Fanuc KAREL source: kt00010.KL

-- PROVISIONAL review KL for V1013-1; original PC SHA256 68f7cc7fb985bd2ba843ab7a48a8a9cfd265290f7bc91fa8e1590b52c63fd289
-- Incomplete behavior may be omitted. Consult companion uncertainty JSON. Do not deploy.
PROGRAM KT00010
%NOLOCKGROUP
VAR
  R1 : REAL
  I2 : INTEGER
  OUT : REAL
BEGIN
  -- UNRESOLVED_PC offsets 5-16; opcodes 2E,23
  -- UNRESOLVED_PC offsets 21-32; opcodes 2E,23
  -- UNRESOLVED_PC offsets 37-57; opcodes 21,21,64,69,23
  -- UNRESOLVED_PC offsets 62-66; opcodes 7F
END KT00010
